// TIA Portal V20 export
// export: Created 2026-11-12T08:00:00.0000000Z, ExportSetting None, DisplayName Totally Integrated Automation Portal, DisplayVersion V20, DisplayName STEP 7 Professional, DisplayVersion V20
FUNCTION_BLOCK "FB_Motor_SealIn_FaultLatch_LAD"   // FB21, LAD
TITLE = FB_Motor_SealIn_FaultLatch_LAD
{ S7_Optimized_Access := 'TRUE' }
// 带故障锁存与防自动重启保护的电机起保停控制（纯LAD实现）
// stored: AutoNumber false, MemoryReserve 10, SetENOAutomatically false
   VAR_INPUT
      startBtn : Bool;
      stopBtn : Bool;
      overloadNC : Bool;
      eStopNC : Bool;
      interlockOk : Bool;
      resetFault : Bool;
   END_VAR
   VAR_OUTPUT
      motorCoil : Bool;
      faultLatched : Bool;
      ready : Bool;
   END_VAR
   VAR
      statRun : Bool;
      statFault : Bool;
   END_VAR
BEGIN

REGION Network 1: 故障置位锁存
   // 网络1：热过载或急停触发时置位锁存故障位
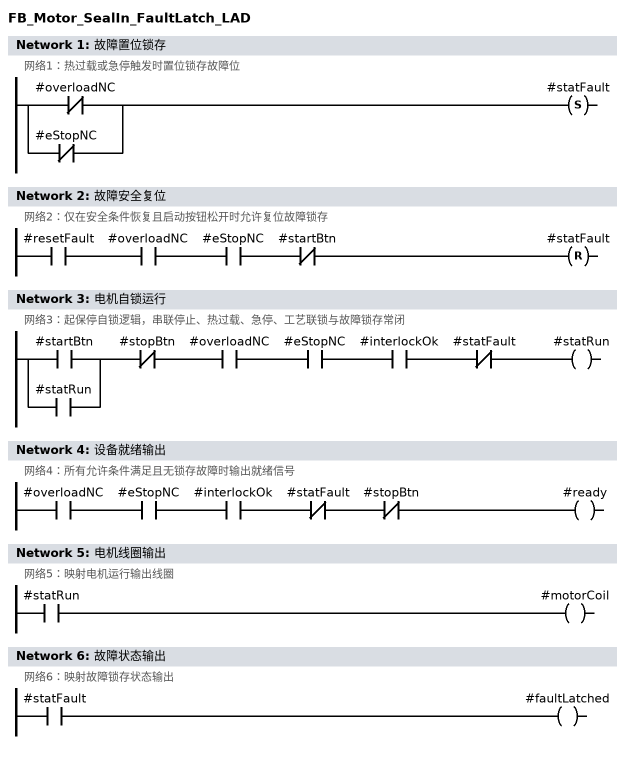
   RUNG wire#powerrail
      I_Contact( #overloadNC )
      wire#w1
      S_Coil( #statFault )
   END_RUNG
   RUNG wire#powerrail
      I_Contact( #eStopNC )
   END_RUNG wire#w1
   // the same network as SCL:
   IF NOT #overloadNC OR NOT #eStopNC THEN #statFault := TRUE; END_IF;
END_REGION

REGION Network 2: 故障安全复位
   // 网络2：仅在安全条件恢复且启动按钮松开时允许复位故障锁存
   RUNG wire#powerrail
      Contact( #resetFault )
      Contact( #overloadNC )
      Contact( #eStopNC )
      I_Contact( #startBtn )
      R_Coil( #statFault )
   END_RUNG
   // the same network as SCL:
   IF #resetFault AND #overloadNC AND #eStopNC AND NOT #startBtn THEN #statFault := FALSE; END_IF;
END_REGION

REGION Network 3: 电机自锁运行
   // 网络3：起保停自锁逻辑，串联停止、热过载、急停、工艺联锁与故障锁存常闭
   RUNG wire#powerrail
      Contact( #startBtn )
      wire#w1
      I_Contact( #stopBtn )
      Contact( #overloadNC )
      Contact( #eStopNC )
      Contact( #interlockOk )
      I_Contact( #statFault )
      Coil( #statRun )
   END_RUNG
   RUNG wire#powerrail
      Contact( #statRun )
   END_RUNG wire#w1
   // the same network as SCL:
   #statRun := (#startBtn OR #statRun) AND NOT #stopBtn AND #overloadNC AND #eStopNC AND #interlockOk AND NOT #statFault;
END_REGION

REGION Network 4: 设备就绪输出
   // 网络4：所有允许条件满足且无锁存故障时输出就绪信号
   RUNG wire#powerrail
      Contact( #overloadNC )
      Contact( #eStopNC )
      Contact( #interlockOk )
      I_Contact( #statFault )
      I_Contact( #stopBtn )
      Coil( #ready )
   END_RUNG
   // the same network as SCL:
   #ready := #overloadNC AND #eStopNC AND #interlockOk AND NOT #statFault AND NOT #stopBtn;
END_REGION

REGION Network 5: 电机线圈输出
   // 网络5：映射电机运行输出线圈
   RUNG wire#powerrail
      Contact( #statRun )
      Coil( #motorCoil )
   END_RUNG
   // the same network as SCL:
   #motorCoil := #statRun;
END_REGION

REGION Network 6: 故障状态输出
   // 网络6：映射故障锁存状态输出
   RUNG wire#powerrail
      Contact( #statFault )
      Coil( #faultLatched )
   END_RUNG
   // the same network as SCL:
   #faultLatched := #statFault;
END_REGION
END_FUNCTION_BLOCK
